(* IEC 61131-3 sources: kns-pump-station/tests/POUs/Log/FB_EventLog_Test, 20 files *)

(* ---- FB_EventLog_Test.decl.st ---- *)
// Назначение: набор coUnit для FB_EventLog — кольцо на 200 записей: запись тревоги и события станции, номер
//             101000 + код, затирание самой старой записи и счётчик, порядок «новые первыми», страницы HMI,
//             курсор внешнего клиента и пропуск затёртых записей, время процесса lrMono_s, снимок для CSV.
//             Журнал (≈16 КБ) — переменная экземпляра метода (VAR_INST), а не стека: тест выполняется
//             за один вызов, повторные вызовы завершённого теста ассерты не проверяют.
// Автор:      kr0nsch
// Версия:     0.1.0
// Документ:   docs/DESIGN.md, разделы 9.1, 14.1
FUNCTION_BLOCK FB_EventLog_Test EXTENDS coUnit.FB_TestSuite
VAR CONSTANT
    LR_EPS_S : LREAL := LREAL#1.0E-6;   // допуск времени процесса, с
    R_EPS : REAL := 1.0E-6;             // допуск значения записи
END_VAR

(* ---- AlarmEventStored.method.decl.st ---- *)
// Событие тревоги: запись вида Alarm со всеми полями события, номер 1, время процесса — по itfTime (1 ч)
METHOD PRIVATE AlarmEventStored
VAR_INST
    fbLog  : FB_EventLog;           // проверяемый журнал
END_VAR
VAR
    fbTime  : PL.FB_FakeTime;       // подменное время, старт 1 ч
    stEvent : PL.ST_AlarmEvent;     // событие тревоги
    stRec   : ST_EventRecord;       // записанная запись
END_VAR

(* ---- EmptyLogDefaults.method.decl.st ---- *)
// Пустой журнал: записей 0, GetRecord — FALSE, одна пустая страница, курсор без строк (первая = последняя + 1)
METHOD PRIVATE EmptyLogDefaults
VAR_INST
    fbLog  : FB_EventLog;           // проверяемый журнал
    stView : ST_EventView;          // страница HMI
    stFeed : ST_EventFeed;          // курсор клиента
END_VAR
VAR
    stRec : ST_EventRecord;         // запись
END_VAR

(* ---- FeedFromSeqOldestFirst.method.decl.st ---- *)
// Курсор: с № 5 — 32 строки № 5…36 от старой к новой; с № 37 — 4 строки и пустые; с № 41 — строк нет
METHOD PRIVATE FeedFromSeqOldestFirst
VAR_INST
    fbLog  : FB_EventLog;           // проверяемый журнал
    stFeed : ST_EventFeed;          // курсор клиента
END_VAR
VAR
    fbTime : PL.FB_FakeTime;        // подменное время
    uiI    : UINT;                  // номер события
END_VAR

(* ---- FeedFromSeqOldestFirst.method.impl.st ---- *)
coUnit.TEST('EventLog_FeedFromSeqOldestFirst');

fbLog.itfTime := fbTime;
FOR uiI := 1 TO 40 DO
    fbLog.LogEvent(eEvent := E_StationEvent.CfgChanged, rValue := UINT_TO_REAL(uiI));
END_FOR
stFeed.udiFromSeq := 5;
fbLog.FillFeed(stFeed := stFeed);
AssertEquals_UINT(Expected := GVL_Const.LOG_FEED_ROWS, Actual := stFeed.uiCount, Message := 'full feed: 32 rows');
AssertEquals_UDINT(Expected := 5, Actual := stFeed.astRow[1].udiSeq, Message := 'row 1 = from');
AssertEquals_UDINT(Expected := 36, Actual := stFeed.astRow[GVL_Const.LOG_FEED_ROWS].udiSeq, Message := 'row 32 = 36');
AssertEquals_UDINT(Expected := 1, Actual := stFeed.udiSeqFirst, Message := 'oldest 1');
AssertEquals_UDINT(Expected := 40, Actual := stFeed.udiSeqLast, Message := 'newest 40');
stFeed.udiFromSeq := 37;
fbLog.FillFeed(stFeed := stFeed);
AssertEquals_UINT(Expected := 4, Actual := stFeed.uiCount, Message := '4 rows from 37');
AssertEquals_UDINT(Expected := 40, Actual := stFeed.astRow[4].udiSeq, Message := 'row 4 = 40');
AssertEquals_UDINT(Expected := 0, Actual := stFeed.astRow[5].udiSeq, Message := 'row 5 cleared');
stFeed.udiFromSeq := 41;
fbLog.FillFeed(stFeed := stFeed);
AssertEquals_UINT(Expected := 0, Actual := stFeed.uiCount, Message := 'nothing new from 41');

coUnit.TEST_FINISHED();

(* ---- FeedReportsOverwrittenGap.method.decl.st ---- *)
// 250 событий: в кольце № 51…250; клиент, ждущий № 10, получает строки с № 51 и видит пропуск по номерам
METHOD PRIVATE FeedReportsOverwrittenGap
VAR_INST
    fbLog  : FB_EventLog;           // проверяемый журнал
    stFeed : ST_EventFeed;          // курсор клиента
END_VAR
VAR
    fbTime : PL.FB_FakeTime;        // подменное время
    uiI    : UINT;                  // номер события
END_VAR

(* ---- FeedReportsOverwrittenGap.method.impl.st ---- *)
coUnit.TEST('EventLog_FeedReportsOverwrittenGap');

fbLog.itfTime := fbTime;
FOR uiI := 1 TO 250 DO
    fbLog.LogEvent(eEvent := E_StationEvent.CfgChanged, rValue := UINT_TO_REAL(uiI));
END_FOR
stFeed.udiFromSeq := 10;
fbLog.FillFeed(stFeed := stFeed);
AssertEquals_UDINT(Expected := 51, Actual := stFeed.udiSeqFirst, Message := 'oldest in ring 51');
AssertEquals_UDINT(Expected := 250, Actual := stFeed.udiSeqLast, Message := 'newest 250');
AssertTrue(Condition := stFeed.udiFromSeq < stFeed.udiSeqFirst, Message := 'client sees gap');
AssertEquals_UDINT(Expected := 51, Actual := stFeed.astRow[1].udiSeq, Message := 'feed starts at oldest');
AssertEquals_UDINT(Expected := 50, Actual := fbLog.udiOverwritten, Message := 'overwritten 50');

coUnit.TEST_FINISHED();

(* ---- GetRecordNewestFirst.method.decl.st ---- *)
// Возраст 0 — самая новая запись; возраст за последней записью — FALSE
METHOD PRIVATE GetRecordNewestFirst
VAR_INST
    fbLog  : FB_EventLog;           // проверяемый журнал
END_VAR
VAR
    fbTime : PL.FB_FakeTime;        // подменное время
    stRec  : ST_EventRecord;        // запись
END_VAR

(* ---- MonoTimeIsProcessTime.method.decl.st ---- *)
// lrMono_s — время процесса по itfTime: разность меток двух записей равна шагу подменных часов (90 с), а не
// настенному времени между вызовами
METHOD PRIVATE MonoTimeIsProcessTime
VAR_INST
    fbLog  : FB_EventLog;           // проверяемый журнал
END_VAR
VAR
    fbTime  : PL.FB_FakeTime;       // подменное время
    stFirst : ST_EventRecord;       // первая запись
    stLast  : ST_EventRecord;       // вторая запись
END_VAR

(* ---- RingOverwritesOldestAndCounts.method.decl.st ---- *)
// 205 событий в кольцо на 200: записей 200, затёрто 5, самая старая — № 6, самая новая — № 205
METHOD PRIVATE RingOverwritesOldestAndCounts
VAR_INST
    fbLog  : FB_EventLog;           // проверяемый журнал
END_VAR
VAR
    fbTime : PL.FB_FakeTime;        // подменное время
    stRec  : ST_EventRecord;        // запись
    uiI    : UINT;                  // номер события
END_VAR

(* ---- RingOverwritesOldestAndCounts.method.impl.st ---- *)
coUnit.TEST('EventLog_RingOverwritesOldestAndCounts');

fbLog.itfTime := fbTime;
FOR uiI := 1 TO 205 DO
    fbLog.LogEvent(eEvent := E_StationEvent.CfgChanged, rValue := UINT_TO_REAL(uiI));
END_FOR
AssertEquals_UINT(Expected := GVL_Const.LOG_CAPACITY, Actual := fbLog.uiCount, Message := 'ring full: 200');
AssertEquals_UDINT(Expected := 5, Actual := fbLog.udiOverwritten, Message := '5 overwritten');
AssertEquals_UDINT(Expected := 205, Actual := fbLog.udiSeqLast, Message := 'last sequence 205');
AssertTrue(Condition := fbLog.GetRecord(uiAge := GVL_Const.LOG_CAPACITY - 1, stRecord => stRec),
           Message := 'oldest present');
AssertEquals_UDINT(Expected := 6, Actual := stRec.udiSeq, Message := 'oldest is no. 6');
AssertEquals_REAL(Expected := 6.0, Actual := stRec.rValue, Delta := R_EPS, Message := 'oldest value 6');
fbLog.GetRecord(uiAge := 0, stRecord => stRec);
AssertEquals_UDINT(Expected := 205, Actual := stRec.udiSeq, Message := 'newest is no. 205');
AssertFalse(Condition := fbLog.GetRecord(uiAge := GVL_Const.LOG_CAPACITY, stRecord => stRec),
            Message := 'no record older than capacity');

coUnit.TEST_FINISHED();

(* ---- SnapshotAfterWrapOldestFirst.method.decl.st ---- *)
// Снимок полного кольца после затирания (205 событий): 200 записей от старой (№ 6) к новой (№ 205) без
// разрыва на границе кольца
METHOD PRIVATE SnapshotAfterWrapOldestFirst
VAR_INST
    fbLog  : FB_EventLog;           // проверяемый журнал
END_VAR
VAR
    fbTime : PL.FB_FakeTime;        // подменное время
    stRec  : ST_EventRecord;        // запись снимка
    uiI    : UINT;                  // номер события и индекс снимка
    uiBad  : UINT;                  // записей снимка не на своём месте
END_VAR

(* ---- SnapshotAfterWrapOldestFirst.method.impl.st ---- *)
coUnit.TEST('EventLog_SnapshotAfterWrapOldestFirst');

fbLog.itfTime := fbTime;
FOR uiI := 1 TO 205 DO
    fbLog.LogEvent(eEvent := E_StationEvent.CfgChanged, rValue := UINT_TO_REAL(uiI));
END_FOR
AssertTrue(Condition := fbLog.TakeSnapshot(), Message := 'snapshot taken');
AssertEquals_UINT(Expected := GVL_Const.LOG_CAPACITY, Actual := fbLog.SnapshotCount, Message := '200 records');
uiBad := 0;
FOR uiI := 0 TO GVL_Const.LOG_CAPACITY - 1 DO
    fbLog.GetSnapshotRecord(uiIndex := uiI, stRecord => stRec);
    IF stRec.udiSeq <> UINT_TO_UDINT(uiI) + 6 THEN
        uiBad := uiBad + 1;
    END_IF
END_FOR
AssertEquals_UINT(Expected := 0, Actual := uiBad, Message := 'index i holds no. i + 6');
fbLog.GetSnapshotRecord(uiIndex := GVL_Const.LOG_CAPACITY - 1, stRecord => stRec);
AssertEquals_UDINT(Expected := 205, Actual := stRec.udiSeq, Message := 'last index newest');

coUnit.TEST_FINISHED();

(* ---- SnapshotIndependentOfLaterEvents.method.decl.st ---- *)
// Снимок — от старой записи к новой; события после снимка его не меняют; индекс вне снимка — FALSE
METHOD PRIVATE SnapshotIndependentOfLaterEvents
VAR_INST
    fbLog  : FB_EventLog;           // проверяемый журнал
END_VAR
VAR
    fbTime : PL.FB_FakeTime;        // подменное время
    stRec  : ST_EventRecord;        // запись снимка
END_VAR

(* ---- StationEventIdIsBasePlusCode.method.decl.st ---- *)
// Событие станции: номер 101000 + код (АВР, код 6 → 101006), вид Station, приоритет None, состояния Normal
METHOD PRIVATE StationEventIdIsBasePlusCode
VAR_INST
    fbLog  : FB_EventLog;           // проверяемый журнал
END_VAR
VAR
    fbTime  : PL.FB_FakeTime;       // подменное время
    itfSink : I_StationEventSink;   // журнал как приёмник событий станции
    stRec   : ST_EventRecord;       // записанная запись
END_VAR

(* ---- TimeBackwardsRecordedAsIs.method.decl.st ---- *)
// «Время назад» (подменные часы с 1 ч на 59 мин 50 с): запись не теряется, номер растёт, метка — как дали часы
METHOD PRIVATE TimeBackwardsRecordedAsIs
VAR_INST
    fbLog  : FB_EventLog;           // проверяемый журнал
END_VAR
VAR
    fbTime : PL.FB_FakeTime;        // подменное время
    stRec  : ST_EventRecord;        // запись
END_VAR

(* ---- ViewPageEqualToCountClamped.method.decl.st ---- *)
// Номер страницы, равный числу страниц (45 записей — страницы 0…2, запрошена 3), — последняя страница (№ 5…1),
// а не пустая страница за концом журнала
METHOD PRIVATE ViewPageEqualToCountClamped
VAR_INST
    fbLog  : FB_EventLog;           // проверяемый журнал
    stView : ST_EventView;          // страница HMI
END_VAR
VAR
    fbTime : PL.FB_FakeTime;        // подменное время
    uiI    : UINT;                  // номер события
END_VAR

(* ---- ViewPageEqualToCountClamped.method.impl.st ---- *)
coUnit.TEST('EventLog_ViewPageEqualToCountClamped');

fbLog.itfTime := fbTime;
FOR uiI := 1 TO 45 DO
    fbLog.LogEvent(eEvent := E_StationEvent.CfgChanged, rValue := UINT_TO_REAL(uiI));
END_FOR
stView.uiPage := 3;
fbLog.FillView(stView := stView);
AssertEquals_UINT(Expected := 2, Actual := stView.uiPage, Message := 'page 3 of 3 clamped to 2');
AssertEquals_UDINT(Expected := 5, Actual := stView.astRow[1].udiSeq, Message := 'last page row 1');

coUnit.TEST_FINISHED();

(* ---- ViewPagination.method.decl.st ---- *)
// 45 записей по 20 строк: 3 страницы; страница 0 — № 45…26, страница 2 — № 5…1 и пустые строки; номер
// страницы больше последней ограничивается последней
METHOD PRIVATE ViewPagination
VAR_INST
    fbLog  : FB_EventLog;           // проверяемый журнал
    stView : ST_EventView;          // страница HMI
END_VAR
VAR
    fbTime : PL.FB_FakeTime;        // подменное время
    uiI    : UINT;                  // номер события
END_VAR

(* ---- ViewPagination.method.impl.st ---- *)
coUnit.TEST('EventLog_ViewPagination');

fbLog.itfTime := fbTime;
FOR uiI := 1 TO 45 DO
    fbLog.LogEvent(eEvent := E_StationEvent.CfgChanged, rValue := UINT_TO_REAL(uiI));
END_FOR
stView.uiPage := 0;
fbLog.FillView(stView := stView);
AssertEquals_UINT(Expected := 3, Actual := stView.uiPageCount, Message := '3 pages');
AssertEquals_UINT(Expected := 45, Actual := stView.uiCount, Message := '45 records');
AssertEquals_UDINT(Expected := 45, Actual := stView.astRow[1].udiSeq, Message := 'page 0 row 1 newest');
AssertEquals_UDINT(Expected := 26, Actual := stView.astRow[GVL_Const.LOG_VIEW_ROWS].udiSeq,
                   Message := 'page 0 last row');
stView.uiPage := 2;
fbLog.FillView(stView := stView);
AssertEquals_UDINT(Expected := 5, Actual := stView.astRow[1].udiSeq, Message := 'page 2 row 1');
AssertEquals_UDINT(Expected := 1, Actual := stView.astRow[5].udiSeq, Message := 'page 2 row 5 oldest');
AssertEquals_UDINT(Expected := 0, Actual := stView.astRow[6].udiSeq, Message := 'page 2 row 6 empty');
stView.uiPage := 7;
fbLog.FillView(stView := stView);
AssertEquals_UINT(Expected := 2, Actual := stView.uiPage, Message := 'page clamped to last');

coUnit.TEST_FINISHED();
